Fanuc KAREL source: kt00265.KL

-- PROVISIONAL review KL for V1013-1; original PC SHA256 08b6cd72949c65cb30255039171e22d81f69d883bb327079c91f855e25b2c263
-- Incomplete behavior may be omitted. Consult companion uncertainty JSON. Do not deploy.
PROGRAM KT00265
%NOLOCKGROUP
VAR
  B1 : BOOLEAN
  B2 : BOOLEAN
  OUT : BOOLEAN
BEGIN
  -- UNRESOLVED_PC offsets 5-12; opcodes 9D,23
  -- UNRESOLVED_PC offsets 17-24; opcodes 9C,23
  -- UNRESOLVED_PC offsets 29-36; opcodes 9D,23
  -- UNRESOLVED_PC offsets 41-48; opcodes 9C,23
  -- UNRESOLVED_PC offsets 53-72; opcodes 21,21,57,23
  -- UNRESOLVED_PC offsets 77-81; opcodes 7F
END KT00265
